(* IEC 61131-3 sources: codesys-framework/txt/application/WeVe General (library)/AirPressure/Hardware/FB_AirPressureHardware, 3 files *)

(* ---- AirPressureOk.prop.st ---- *)
PROPERTY AirPressureOk : BOOL

// --- BEGIN IMPLEMENTATION ---

// ----------- GET -----------
VAR
	scSignals 	: SC_DigitalInputSignals;
END_VAR

// -- BEGIN IMPLEMENTATION GET --
scSignals := _fbAirPressure.Signals;

AirPressureOk := scSignals.xDIDelayedDetectionStateOff;

(* ---- LoadHardCodedSettings.method.st ---- *)
METHOD PROTECTED LoadHardCodedSettings
VAR_INPUT
END_VAR

// --- BEGIN IMPLEMENTATION ---

_scSysParAirPressure.eSysPar_DI_SensorType := E_DigitalInputSensorType.Type_NO;
_scSysParAirPressure.tSysPar_Detection_OnDelay := T#1S;
_scSysParAirPressure.tSysPar_Detection_OffDelay := T#1S;
_scSysParAirPressure.tSysPar_Detection_OnDelayOnOff := T#1S;
_scSysParAirPressure.tSysPar_Detection_OffDelayOnOff := T#1S;

(* ---- ProcessHardware.method.st ---- *)
METHOD PROTECTED ProcessHardware
VAR_INPUT
END_VAR

// --- BEGIN IMPLEMENTATION ---

_fbAirPressure.SysPar := _scSysParAirPressure;
_fbAirPressure();
